Fanuc KAREL source: kf00116.KL

-- PROVISIONAL review KL for V940-1; original PC SHA256 d46327ea168f10c96727ba4f24f85ba3ed1e1dede43fc605501404419b0f7dec
-- Incomplete behavior may be omitted. Consult companion uncertainty JSON. Do not deploy.
PROGRAM KF00116
%NOLOCKGROUP
BEGIN
  -- V9_EXPOSED_INDEXED_TABLE_HINT layout=0001; 2 counted words exposed once; source arms/runtime held
  -- UNRESOLVED_PC offsets 0-1; opcodes 7B
  -- UNRESOLVED_PC offsets 6-19; opcodes 2D,9D,5A,79
  -- UNRESOLVED_PC offsets 24-29; opcodes 9D,7F
  -- UNRESOLVED_PC offsets 34-39; opcodes 7A
  -- UNRESOLVED_PC offsets 44-68; opcodes 2D,27,27,2D,9D,53,AA,54,7F
  -- UNRESOLVED_PC offsets 78-82; opcodes 7F
  -- UNRESOLVED_PC offsets 87-103; opcodes 27,27,2E,AA,23
  -- UNRESOLVED_PC offsets 108-112; opcodes 7F
END KF00116
